// TIA Portal V21 export
// export: Created 2026-11-03T19:44:49.7617988Z, ExportSetting WithDefaults, WithReadOnly, DisplayName Totally Integrated Automation Portal, DisplayVersion V21, DisplayName STEP 7 Professional, DisplayVersion V21, DisplayName STEP 7 Safety, DisplayVersion V21, DisplayName Tech WebApplication, DisplayVersion V21, DisplayName WinCC Basic/Comfort/Advanced, DisplayVersion V21, DisplayName WinCC Professional, DisplayVersion V21, DisplayName WinCC Unified, DisplayVersion V21
ORGANIZATION_BLOCK "Main"   // OB1, SCL, ProgramCycle
{ S7_Optimized_Access := 'TRUE' }
VERSION : 1.0
// SPDX-License-Identifier: MIT. No equipment library or process sequence.
// stored: AutoNumber true, CodeModifiedDate 2026-11-03T19:44:43.8400479Z, CompileDate 2026-11-03T19:44:43.8400479Z, ConstantName OB_Main, CreationDate 2026-11-03T19:44:33.7000652Z, DownloadDate 0001-01-01T00:00:00Z, EventClass Program cycle, HandleErrorsWithinBlock false, InterfaceModifiedDate 2026-11-03T19:44:33.988557Z, IsConsistent true, IsIECCheckEnabled false, IsKnowHowProtected false, IsWriteProtected false, LoadMemoryLength 14729, ModifiedDate 2026-11-03T19:44:43.8400479Z, PLCSimAdvancedSupport true, ParameterModified 2026-11-03T19:44:33.9885569Z, PriorityNumber 1, ProcessImagePartNumber 65535, SetENOAutomatically false, StructureModified 2026-11-03T19:44:33.988557Z, VirtualPlcSupport false, WorkMemoryLength 554
   VAR_INPUT
      Initial_Call : Bool;   // Initial call of this OB
      Remanence : Bool;   // =True, if remanent data are available
   END_VAR
BEGIN

       "DB_FAT_Demo".P101_RunCommand := "DB_FAT_Demo".EnableDemo AND "DB_FAT_Demo".StopHealthy AND "DB_FAT_Demo".P101_Request;
       IF "DB_FAT_Demo".P101_RunCommand THEN
           "DB_FAT_Demo".P101_SpeedCommand := LIMIT(MN := REAL#0.0, IN := "DB_FAT_Demo".P101_RequestedSpeed, MX := REAL#100.0);
       ELSE
           "DB_FAT_Demo".P101_SpeedCommand := REAL#0.0;
       END_IF;
       "DB_FAT_Demo".P201_RunCommand := "DB_FAT_Demo".EnableDemo AND "DB_FAT_Demo".StopHealthy AND "DB_FAT_Demo".P201_Request;
       IF "DB_FAT_Demo".P201_RunCommand THEN
           "DB_FAT_Demo".P201_SpeedCommand := LIMIT(MN := REAL#0.0, IN := "DB_FAT_Demo".P201_RequestedSpeed, MX := REAL#100.0);
       ELSE
           "DB_FAT_Demo".P201_SpeedCommand := REAL#0.0;
       END_IF;
       "DB_FAT_Demo".P202_RunCommand := "DB_FAT_Demo".EnableDemo AND "DB_FAT_Demo".StopHealthy AND "DB_FAT_Demo".P202_Request;
       IF "DB_FAT_Demo".P202_RunCommand THEN
           "DB_FAT_Demo".P202_SpeedCommand := LIMIT(MN := REAL#0.0, IN := "DB_FAT_Demo".P202_RequestedSpeed, MX := REAL#100.0);
       ELSE
           "DB_FAT_Demo".P202_SpeedCommand := REAL#0.0;
       END_IF;
       "DB_FAT_Demo".P301_RunCommand := "DB_FAT_Demo".EnableDemo AND "DB_FAT_Demo".StopHealthy AND "DB_FAT_Demo".P301_Request;
       IF "DB_FAT_Demo".P301_RunCommand THEN
           "DB_FAT_Demo".P301_SpeedCommand := LIMIT(MN := REAL#0.0, IN := "DB_FAT_Demo".P301_RequestedSpeed, MX := REAL#100.0);
       ELSE
           "DB_FAT_Demo".P301_SpeedCommand := REAL#0.0;
       END_IF;
       "DB_FAT_Demo".XV101_OpenCommand := "DB_FAT_Demo".EnableDemo AND "DB_FAT_Demo".StopHealthy AND "DB_FAT_Demo".XV101_Request;
       "DB_FAT_Demo".XV201_OpenCommand := "DB_FAT_Demo".EnableDemo AND "DB_FAT_Demo".StopHealthy AND "DB_FAT_Demo".XV201_Request;
       "DB_FAT_Demo".XV202_OpenCommand := "DB_FAT_Demo".EnableDemo AND "DB_FAT_Demo".StopHealthy AND "DB_FAT_Demo".XV202_Request;
       "DB_FAT_Demo".XV301_OpenCommand := "DB_FAT_Demo".EnableDemo AND "DB_FAT_Demo".StopHealthy AND "DB_FAT_Demo".XV301_Request;
       "DB_FAT_Demo".XV102_OpenCommand := "DB_FAT_Demo".EnableDemo AND "DB_FAT_Demo".StopHealthy AND "DB_FAT_Demo".XV102_Request;
       "DB_FAT_Demo".XV203_OpenCommand := "DB_FAT_Demo".EnableDemo AND "DB_FAT_Demo".StopHealthy AND "DB_FAT_Demo".XV203_Request;
       "DB_FAT_Demo".XV103_OpenCommand := "DB_FAT_Demo".EnableDemo AND "DB_FAT_Demo".StopHealthy AND "DB_FAT_Demo".XV103_Request;
       IF "DB_FAT_Demo".EnableDemo AND "DB_FAT_Demo".StopHealthy THEN
           "DB_FAT_Demo".FCV302_PositionCommand := LIMIT(MN := REAL#0.0, IN := "DB_FAT_Demo".FCV302_RequestedPosition, MX := REAL#100.0);
       ELSE
           "DB_FAT_Demo".FCV302_PositionCommand := REAL#0.0;
       END_IF;
       "DB_FAT_Demo".LT101_Percent := SCALE_X(MIN := REAL#0.0,
           VALUE := NORM_X(MIN := INT#0, VALUE := "DB_FAT_Demo".LT101_Raw, MAX := INT#27648), MAX := REAL#100.0);
       "DB_FAT_Demo".LT201_Percent := SCALE_X(MIN := REAL#0.0,
           VALUE := NORM_X(MIN := INT#0, VALUE := "DB_FAT_Demo".LT201_Raw, MAX := INT#27648), MAX := REAL#100.0);
       "DB_FAT_Demo".LT301_Percent := SCALE_X(MIN := REAL#0.0,
           VALUE := NORM_X(MIN := INT#0, VALUE := "DB_FAT_Demo".LT301_Raw, MAX := INT#27648), MAX := REAL#100.0);
END_ORGANIZATION_BLOCK
